{attribute 'qualified_only'}
{attribute 'strict'}
{attribute 'to_string'}
TYPE E_UDint :
(
	eOptionA := 0,
	eOptionB,
	eOptionC
) UDINT;
END_TYPE

(* stored: Version 1.1.0.1, ProductVersion 3.1.4026.19
   DUT E_UDint: Id {2b5f7952-8b04-4766-8791-9b0549c8c7bc} *)
